// TIA Portal V18 export
TYPE "TargetProductionMdz_in"
   STRUCT
      KPI_Informations : Struct
         Full_AvailabilityShift : Array[1.."ShiftList_Setup_Const"] of Time;
         Full_AvailabilityDay : Time := T#9H_15M;
         Net_AvailabilityShift : Array[1.."ShiftList_Setup_Const"] of Time;
         Net_AvailabilityDay : Time := T#9H_15M;
         Total_StopPlannedShift : Array[1.."ShiftList_Setup_Const"] of Time;
         Total_StopPlannedDay : Time := T#0MS;
         StopPlanned_Executed_Shift : Array[1.."ShiftList_Setup_Const"] of Time;
         StopPlanned_Executed_Day : Time := T#2H_45M;
         NextStopPlanned : Date_And_Time := DT#2000-01-10-00:00:00;
         NextStopPlanned_Index : Int := 11;
         RemaningTimeToStopPlanned : Time := T#8D_15H_45M_48S_109MS;
         NextStopPlannedInRealTime : Time := T#8H_14M_11S_891MS;
         RemaningCycleToStoPplanned : DInt := 2_139_095_040;
         Total_StopTimeShift : Array[1.."ShiftList_Setup_Const"] of Time;
         Total_StopTimeDay : Time := T#-1H_41M_28S;
         GoalOfShift : Array[1.."ShiftList_Setup_Const"] of Int;
         GoalOfDay : Int := 199;
         TaktStandardByShift : Array[1.."ShiftList_Setup_Const"] of Time;
      END_STRUCT;
      KPI_Results : Struct
         Production_Status : Int := 0;
         MaxProductionCapacity_Shift : Array[1.."ShiftList_Setup_Const"] of Int;
         MaxProductionCapacity_Day : Int := 246;
         TimeToProductionDone_Shift : Array[1.."ShiftList_Setup_Const"] of Time;
         TimeToProductionDone_Day : Time := T#0MS;
      END_STRUCT;
   END_STRUCT;
   // KPI_Informations.Full_AvailabilityShift[1] := T#9H_15M;
   // KPI_Informations.Full_AvailabilityShift[2..3] := T#0MS;
   // KPI_Informations.Net_AvailabilityShift[1] := T#9H_15M;
   // KPI_Informations.Net_AvailabilityShift[2..3] := T#0MS;
   // KPI_Informations.Total_StopPlannedShift[1..3] := T#0MS;
   // KPI_Informations.StopPlanned_Executed_Shift[1] := T#1H_35M;
   // KPI_Informations.StopPlanned_Executed_Shift[2] := T#1H_10M;
   // KPI_Informations.StopPlanned_Executed_Shift[3] := T#0MS;
   // KPI_Informations.Total_StopTimeShift[1] := T#-1H_11M_58S;
   // KPI_Informations.Total_StopTimeShift[2] := T#-29M_30S;
   // KPI_Informations.Total_StopTimeShift[3] := T#0MS;
   // KPI_Informations.GoalOfShift[1] := 164;
   // KPI_Informations.GoalOfShift[2] := 35;
   // KPI_Informations.GoalOfShift[3] := 0;
   // KPI_Informations.TaktStandardByShift[1] := T#2M_15S;
   // KPI_Informations.TaktStandardByShift[2] := T#10M;
   // KPI_Informations.TaktStandardByShift[3] := T#0MS;
   // KPI_Results.MaxProductionCapacity_Shift[1] := 246;
   // KPI_Results.MaxProductionCapacity_Shift[2..3] := 0;
   // KPI_Results.TimeToProductionDone_Shift[1..3] := T#0MS;
END_TYPE
